INTERFACE iLightCmdSource

METHOD Process
VAR_IN_OUT
	CmdEvent : stLightCmdEvent;
END_VAR
END_METHOD

END_INTERFACE

(* stored: Version 1.1.0.1
   Itf iLightCmdSource: Id {dbabc1f4-79bd-44f7-9985-dadc5324c1ab}
   Method Process: Id {020f83b5-ca73-4be5-8db2-53f02b4a1991} *)
